{attribute 'qualified_only'}
TYPE E_AnalogInputCommand : (NONE := 0, MEASURE := 1) DINT;
END_TYPE

(* stored: Version 1.1.0.1, ProductVersion 3.1.4024.12
   DUT E_AnalogInputCommand: Id {0acb6598-db4f-4461-bd02-ebe85f2f8009} *)
